TYPE ST_PwmOutput_HMI EXTENDS ST_HmiFunction :
	STRUCT
		// Commands from the HMI (only applied while the HMI function is enabled)
		RpmSetpoint		  : LREAL; // [rpm]
		FrequencySetpoint : LREAL := 100; // [Hz]
		Reset			  : BOOL;  // Acknowledge PWM error, cleared by the PLC
		// Status to the HMI
		Rpm				  : LREAL; // [rpm] actual, calculated back from the duty cycle
		DutyCycle		  : LREAL; // [%]
		Frequency		  : LREAL := 100; // [Hz]
		Error			  : BOOL;
		Warning			  : BOOL;
	END_STRUCT
END_TYPE

(* stored: Version 1.1.0.1
   DUT ST_PwmOutput_HMI: Id {66fbf164-0150-4285-a7aa-fceaba346305} *)
